(* IEC 61131-3 sources: daoli-st-library/DL_Process (part 60) *)

(* ---- FB_DL_AgvDockingHandshake.st ---- *)
(*==============================================================================
 * 组件名称 (Component)  : FB_DL_AgvDockingHandshake
 * 所属子库 (Sublibrary) : DL_Process
 * 当前版本 (Version)    : 1.0.1
 * 组件分类 (Category)   : 功能块（FUNCTION_BLOCK）· 工站模板 · 移动载体对接交接
 * 兼容性 (Platform)     : CODESYS 3.5 / TwinCAT 3 / 汇川 InoProShop / Machine Expert；
 *                         仅依赖标准库（TON / R_TRIG / F_TRIG），握手信号全部为布尔
 *                         引脚注入，块内不含任何车辆调度、导航或总线通讯细节
 * 功能描述 (Function)   : 把「到位检测 → 双侧就绪握手 → 交接放行 → 完成确认」做成带
 *                         超时与失序诊断的交接状态机，屏蔽移动载体与固定工站两侧的
 *                         信号时序差异，产出单一放行位与握手成功单拍脉冲
 * 与既有件边界 (Scope)  : 固定段之间的连续物流握手（成组上下游节拍链）由输送链路件
 *                         承担，属长连接；本件面向移动载体与固定工站的临时对接（会话
 *                         式、一次性），握手条件含「物料在位」与「双侧就绪」双约束，
 *                         语义与生命周期都不同，不可互替
 * 状态机规模 (States)   : 七态（eIdle 0 / eWaitArrive 10 / eDockConfirm 20 /
 *                         ePermitTransfer 30 / eTransferMonitor 40 / eComplete 50 /
 *                         eFault 99）；编号留 10 间隔便于插态
 * 关键算法 (Algorithm)  :
 *   ① 到位稳定：到位信号须连续两个扫描周期为真才推进，滤掉光电单拍毛刺
 *   ② 双侧就绪：两侧就绪位须同时为真且连续两拍成立，避免单拍毛刺直接放行
 *   ③ 物料一致性：进入交接监视时快照物料在位位；过程中该位由真转假且完成确认尚未
 *      到达，即判物料丢失或错位（02E2），因为这属于「该在的时候不在」
 *   ④ 完成判定：完成确认上升沿 → 置完成保持位、对接次数累加、撤放行、出握手单拍
 *   ⑤ 失序诊断：完成确认在到位或握手阶段提前到达，属非法请求序列（02E3），直接锁
 *      故障而不吞掉，否则上游误接线会被解释成「一次成功交接」
 *   ⑥ 状态停留时长：用「状态未变则计时、状态一变即清零」的单一秒表实现，供现场
 *      判读卡在哪个阶段，不额外增加引脚
 * 码位表 (Error codes)  :
 *   16#0005_01C3【信息级】超时参数越界已钳位，不置故障位
 *   16#0005_02E0【故障级】到位确认超时
 *   16#0005_02E1【故障级】握手或交接超时（两处共用，均属未在期望时间内建立期望状态）
 *   16#0005_02E2【故障级】物料在位信号丢失
 *   16#0005_02E3【故障级】非法请求序列（完成确认提前到达）
 *   16#0005_02E4【故障级】非法状态兜底
 * R32 写入点次序审计 :
 *   bTransferComplete : ① 待机启动拍清（eIdle）→ ② 交接监视完成拍置（eTransferMonitor
 *                       ，唯一置位点）。保持特性由「不再写」实现，不设第三处写点
 *   _uErrorIdInt      : ① 首扫清（段 4）→ ② 到位超时（eWaitArrive）→ ③ 握手/交接超时
 *                       （eDockConfirm 与 eTransferMonitor 各一处，同拍只命中一处）
 *                       → ④ 物料丢失（eTransferMonitor）→ ⑤ 失序（段 5）→ ⑥ 非法状态
 *                       （ELSE）→ ⑦ 复位清（eFault）
 *   _eState           : 每拍只在 CASE 分支出口单点写入；CASE 之外仅两处（段 5 失序监视、
 *                       段 6 中止与使能撤销），均在 CASE 之前，次序固定
 *   _bMatSnap         : ① 交接监视入口快照（ePermitTransfer 转出拍）→ ② 完成与复位清
 *   tElapsed          : 仅段 10 单点派生（秒表已历时），状态机内不写
 * 设计偏离登记 (Deviations) :
 *   D1 bHandshakeOk 取「握手成功」口径，在进入放行态那一拍出脉冲；规格验收向量 V1 把
 *      该脉冲写在完成确认之后叙述，二者不冲突——脉冲发生在交接放行时刻，完成确认只
 *      负责置完成保持位，头注释按状态迁移表口径落地
 *   D2 到位与双侧就绪用「连续两拍」替代「沿后与门」等价实现，效果相同（滤单拍毛刺），
 *      但不需要额外的边沿实例，拍序更易推演
 * 验收向量 (Acceptance) :
 *   V1 正常序：到位 → 双侧就绪依序为真 → 放行位为真、握手单拍、完成确认后完成保持位
 *      为真且对接次数加一
 *   V2 到位超时：超时窗 10 秒内到位信号未建立 → 码 02E0、故障态
 *   V3 物料丢失：交接监视内物料在位由真转假且完成确认为假 → 码 02E2、放行位撤
 *   V4 完成提前：到位阶段完成确认为真 → 码 02E3、直接故障态
 *   V5 统计：交接监视停留 12 秒、监视超时 30 秒 → 上一轮时长 12 秒、累计加 12 秒
 * 开源溯源 (Origin)     : 参考包装机械与批控公开手册的「会话式交接」阶段划分与双侧
 *                         就绪语义组织，只借阶段分类与参数域；状态机、快照一致性判据、
 *                         失序诊断、码位与引脚契约为本库独立设计，clean-room 不构成
 *                         衍生作品
 * 红线自检 (Redline)    : R1 零全局表与外部变量引用、零物理地址记号 ✓｜R2 零占位符 ✓
 *                         R3 纯 IEC 61131-3 加标准库 ✓｜R4 时长比较带零值旁路、计数
 *                         饱和、无数组访问 ✓｜R5 声明行中英双语同行注释 ✓｜R6 七成员
 *                         逐一有 CASE 标签且含 ELSE 兜底 ✓｜R7 三沿检测与四定时器全
 *                         部在 CASE 之外无条件刷新 ✓
 * 修订历史 (Revision)   :
 *   2026-11-15  v1.0.0  首版入库（Round 11 · C 泳道 · 工站四件套之三）
 *   2026-11-16  v1.0.1  R13 机检 R39 修复：段 5 使能撤销分支原先把 _eState 无条件
 *                       改写为 eIdle，而故障复位沿的消化位于其后 CASE 的 eFault
 *                       分支——禁用期间按下的复位沿当拍被抹掉，_bFaultLatch 与
 *                       故障码留存至操作员补按第二次复位，期间使能回升也被
 *                       「有锁存」判据挡在待机。改为 eFault 态不被禁用覆盖
 *============================================================================*)

(*------------------------------------------------------------------------------
 * 枚举: E_DL_AgvDockState（归属 FB_DL_AgvDockingHandshake，同文件发布）
 *   七态，每个成员在主状态机中均有同名 CASE 标签（R31 完备性）
 *-----------------------------------------------------------------------------*)
TYPE E_DL_AgvDockState :
(
    eIdle            := 0,  // 待机：等到位信号 / Idle, awaiting arrival signal
    eWaitArrive      := 10, // 到位确认：等到位信号稳定 / Arrival confirmation, waiting for a stable signal
    eDockConfirm     := 20, // 对接确认：等双侧就绪同时成立 / Dock confirmation, waiting for both sides ready
    ePermitTransfer  := 30, // 放行交接：单拍过渡态 / Transfer permit, a single-scan transition state
    eTransferMonitor := 40, // 交接监视：等完成确认并监视物料在位 / Transfer monitor, watching completion and material
    eComplete        := 50, // 交接完成：保持一拍后回待机 / Complete, holds one scan then returns
    eFault           := 99  // 故障锁存：仅复位沿可退 / Fault latched, only a reset edge leaves
);
END_TYPE

(*------------------------------------------------------------------------------
 * 结构体: ST_DL_AgvDockStat（归属 FB_DL_AgvDockingHandshake）
 *   跨周期统计，由调用方持有，本块只累加，掉电保持由上层负责
 *-----------------------------------------------------------------------------*)
TYPE ST_DL_AgvDockStat :
STRUCT
    nDockCount     : UDINT;                 // 累计成功对接次数 [次] [Docking counter]
    tTotalTransfer : TIME;                  // 累计交接时长 [毫秒] [Accumulated transfer time]
    tLastCycle     : TIME;                  // 上一轮交接时长 [毫秒] [Last transfer duration]
END_STRUCT
END_TYPE

FUNCTION_BLOCK FB_DL_AgvDockingHandshake
VAR_INPUT
    bEnable           : BOOL;               // 使能，FALSE 撤回全部放行位 [Enable, withdraws all permits on FALSE]
    bReset            : BOOL;               // 复位故障，上升沿受理 [Reset fault on rising edge]
    bAbort            : BOOL;               // 中止本次交接，上升沿受理，不置故障 [Abort the handshake on rising edge, no fault]
    bAgvArrived       : BOOL;               // 载体到位光电（粗定位）[-] [Carrier presence sensor]
    bAgvDockReady     : BOOL;               // 载体侧对接机构就绪 [-] [Carrier-side dock ready]
    bStationReady     : BOOL;               // 工站侧可收料或可放料 [-] [Station-side ready]
    bMaterialOnAgv    : BOOL;               // 物料在位，交接前为载侧、交接后为站侧 [-] [Material present flag]
    bTransferDone     : BOOL;               // 下游完成接收确认 [-] [Downstream receipt confirmation]
    tArriveTimeout    : TIME := T#10S;      // 到位确认超时 [毫秒]，0 表示不监控 [Arrival timeout]
    tHandshakeTimeout : TIME := T#5S;       // 双侧就绪握手超时 [毫秒]，0 表示不监控 [Handshake timeout]
    tTransferTimeout  : TIME := T#30S;      // 交接过程超时 [毫秒]，0 表示不监控 [Transfer timeout]
END_VAR
VAR_OUTPUT
    bDockLamp         : BOOL;               // 对接允许指示灯，载体可进入 [-] [Dock-permitted lamp]
    bTransferPermit   : BOOL;               // 放行交接，可放料或可接料 [-] [Transfer permit]
    bHandshakeOk      : BOOL;               // 握手成功单拍脉冲 [-] [Single pulse when handshake succeeds]
    bTransferComplete : BOOL;               // 交接完成，保持到下次启动 [Transfer complete, held until next cycle]
    eState            : E_DL_AgvDockState;  // 主状态机当前态 [-] [Current state]
    bError            : BOOL;               // 故障锁存，需复位清除 [Latched fault]
    uErrorId          : UDINT;              // 事件码或故障码，0 表示无 [Event or fault code]
    tElapsed          : TIME;               // 当前态已耗时 [毫秒]，现场判读用 [Elapsed time in current state]
END_VAR
VAR_IN_OUT
    stStat            : ST_DL_AgvDockStat;  // 跨周期统计，调用方持有 [Persistent statistics]
END_VAR
VAR
    _eState          : E_DL_AgvDockState := E_DL_AgvDockState.eIdle;  // 内部状态寄存器，唯一真值源 [Internal state register]
    _eStateIn        : E_DL_AgvDockState := E_DL_AgvDockState.eIdle;  // 上拍状态，用于识别迁移拍 [Previous state of last scan]
    _bInit           : BOOL := FALSE;       // 首扫标志，初值 FALSE，判据 NOT _bInit [First-scan flag, R19 pattern]
    _bFaultLatch     : BOOL;                // 故障级锁存，仅复位路径清 [Fault latch, reset path only]
    _uErrorIdInt     : UDINT;               // 故障级码寄存 [Fault-level code register]
    _uInfoCode       : UDINT;               // 本拍信息级码，每拍重算 [Transient info code]
    _bStateChg       : BOOL;                // 本拍发生过状态迁移，秒表清零用 [State changed this scan]
    _bArrivePrev     : BOOL;                // 上位到位信号，稳定判据用 [Arrival signal of last scan]
    _bBothReadyPrev  : BOOL;                // 上拍双侧就绪，稳定判据用 [Both-ready of last scan]
    _bMatSnap        : BOOL;                // 交接入口物料在位快照 [Material snapshot at monitor entry]
    tArriveEff       : TIME;                // 生效到位超时 [毫秒] [Effective arrival timeout]
    tHandEff         : TIME;                // 生效握手超时 [毫秒] [Effective handshake timeout]
    tTranEff         : TIME;                // 生效交接超时 [毫秒] [Effective transfer timeout]
    tMoniEff         : TIME;                // 本次交接监视时长（钳位后）[毫秒] [Clamped monitor duration]
    bArriveIn        : BOOL;                // 到位计时输入条件，先算后调 [Arrival timer input]
    bHandIn          : BOOL;                // 握手计时输入条件，先算后调 [Handshake timer input]
    bTranIn          : BOOL;                // 交接计时输入条件，先算后调 [Transfer timer input]
    fbTrigReset      : R_TRIG;              // 复位沿检测 [Reset edge detector]
    fbTrigAbort      : R_TRIG;              // 中止沿检测 [Abort edge detector]
    fbTrigDone       : R_TRIG;              // 完成确认上升沿 [Completion rising edge]
    fbTrigMateria    : F_TRIG;              // 物料在位下降沿，丢失诊断用 [Material falling edge, loss diagnosis]
    fbTmoArrive      : TON;                 // 到位确认计时 [Arrival timer]
    fbTmoHandshake   : TON;                 // 双侧就绪握手计时 [Handshake timer]
    fbTmoTransfer    : TON;                 // 交接过程计时 [Transfer timer]
    fbTmoState       : TON;                 // 状态停留秒表 [State elapsed stopwatch]
END_VAR
VAR CONSTANT
    DL_FLOAT_EPS     : REAL := 1.0E-6;      // 浮点判等容差（预留）[-] [Float comparison epsilon]
    DL_STAT_MAX      : UDINT := 16#FFFF_FFFE; // 统计计数饱和上限 [次] [Statistics saturation limit]
    DL_TMO_MAX       : TIME := T#600S;      // 超时参数域上限 [毫秒] [Timeout upper bound]
    DL_TMAX_STATE    : TIME := T#24H;       // 状态秒表量程 [毫秒] [State stopwatch range]
    DL_TIME_MAX      : TIME := T#500H;     // 累计时长饱和上限 [毫秒] [Duration saturation limit]
    DL_INFO_TMO_CLAMP: UDINT := 16#0005_01C3; // 01C3 超时参数越界已钳位【信息级】 [Info, timeout clamped]
    DL_ERR_ARRIVE    : UDINT := 16#0005_02E0; // 02E0 到位确认超时【故障级】 [Fault, arrival timeout]
    DL_ERR_HANDSHAKE : UDINT := 16#0005_02E1; // 02E1 握手或交接超时【故障级】 [Fault, handshake or transfer timeout]
    DL_ERR_MATERIAL  : UDINT := 16#0005_02E2; // 02E2 物料在位信号丢失【故障级】 [Fault, material lost]
    DL_ERR_SEQUENCE  : UDINT := 16#0005_02E3; // 02E3 非法请求序列【故障级】 [Fault, illegal request sequence]
    DL_ERR_STATE     : UDINT := 16#0005_02E4; // 02E4 非法状态兜底【故障级】 [Fault, illegal state]
END_VAR

// ==== 段 1｜单拍输出预清零（握手脉冲每拍先清零，置位点唯一） / Single-scan pulse pre-clear, single set point
bHandshakeOk := FALSE;                      // 握手单拍先清零 [Handshake pulse pre-cleared]
_uInfoCode   := 16#0000_0000;               // 信息级码每拍重算 [Info code recomputed]

// ==== 段 2｜超时参数钳位（三个超时统一钳位，零值表示不监控） / Timeout clamping, zero disables supervision
tArriveEff := tArriveTimeout;               // 到位超时先取引脚值 [Arrival timeout from pin]
IF tArriveEff > DL_TMO_MAX THEN
    tArriveEff := DL_TMO_MAX;               // 超上限钳位 [Clamped to upper bound]
    _uInfoCode := DL_INFO_TMO_CLAMP;        // 01C3 超时参数越界已钳位【信息级】 [Info, timeout clamped]
ELSIF tArriveEff < T#0S THEN
    tArriveEff := T#0S;                     // 负值归零即不监控 [Negative means disabled]
END_IF

tHandEff := tHandshakeTimeout;              // 握手超时先取引脚值 [Handshake timeout from pin]
IF tHandEff > DL_TMO_MAX THEN
    tHandEff   := DL_TMO_MAX;               // 超上限钳位 [Clamped to upper bound]
    _uInfoCode := DL_INFO_TMO_CLAMP;        // 01C3 超时参数越界已钳位【信息级】 [Info, timeout clamped]
ELSIF tHandEff < T#0S THEN
    tHandEff := T#0S;                       // 负值归零即不监控 [Negative means disabled]
END_IF

tTranEff := tTransferTimeout;               // 交接超时先取引脚值 [Transfer timeout from pin]
IF tTranEff > DL_TMO_MAX THEN
    tTranEff   := DL_TMO_MAX;               // 超上限钳位 [Clamped to upper bound]
    _uInfoCode := DL_INFO_TMO_CLAMP;        // 01C3 超时参数越界已钳位【信息级】 [Info, timeout clamped]
ELSIF tTranEff < T#0S THEN
    tTranEff := T#0S;                       // 负值归零即不监控 [Negative means disabled]
END_IF

// ==== 段 3｜沿与定时器无条件刷新（R7 红线：严禁置于 IF / CASE 分支内） / Unconditional refresh of edges and timers
fbTrigReset(CLK := bReset);                 // 复位沿 [Reset edge]
fbTrigAbort(CLK := bAbort);                 // 中止沿 [Abort edge]
fbTrigDone(CLK := bTransferDone);           // 完成确认上升沿 [Completion rising edge]
fbTrigMateria(CLK := bMaterialOnAgv);       // 物料在位下降沿 [Material falling edge]

IF (_eState = E_DL_AgvDockState.eWaitArrive) AND (tArriveEff > T#0S) THEN
    bArriveIn := TRUE;                      // 仅到位段且监控开启时计时 [Only while waiting with supervision on]
ELSE
    bArriveIn := FALSE;                     // 其余段清零 [Cleared otherwise]
END_IF
fbTmoArrive(IN := bArriveIn, PT := tArriveEff);

IF (_eState = E_DL_AgvDockState.eDockConfirm) AND (tHandEff > T#0S) THEN
    bHandIn := TRUE;                        // 仅握手段且监控开启时计时 [Only while confirming with supervision on]
ELSE
    bHandIn := FALSE;                       // 其余段清零 [Cleared otherwise]
END_IF
fbTmoHandshake(IN := bHandIn, PT := tHandEff);

IF (_eState = E_DL_AgvDockState.eTransferMonitor) AND (tTranEff > T#0S) THEN
    bTranIn := TRUE;                        // 仅交接段且监控开启时计时 [Only while monitoring with supervision on]
ELSE
    bTranIn := FALSE;                       // 其余段清零 [Cleared otherwise]
END_IF
fbTmoTransfer(IN := bTranIn, PT := tTranEff);

// 状态秒表：本拍未发生迁移才计时；迁移后的下一拍输入断一拍，已历时清零（时基由定时器内部保证）
fbTmoState(IN := (NOT _bStateChg) AND bEnable, PT := DL_TMAX_STATE);

// ==== 段 4｜首扫初始化（R19 唯一合法范式：初值 FALSE，判据 NOT，同步后置 TRUE） / First-scan initialisation with the canonical R19 pattern
IF NOT _bInit THEN
    _eState          := E_DL_AgvDockState.eIdle;  // 状态回待机 [State to idle]
    _eStateIn        := E_DL_AgvDockState.eIdle;  // 上拍状态同步 [Previous state synced]
    _bFaultLatch     := FALSE;              // 故障锁存清零 [Fault latch cleared]
    _uErrorIdInt     := 16#0000_0000;       // 故障码清零 [Fault code cleared]
    _bStateChg       := FALSE;              // 迁移标志清零 [State change flag cleared]
    _bArrivePrev     := FALSE;              // 到位上拍值清零 [Arrival previous cleared]
    _bBothReadyPrev  := FALSE;              // 双侧就绪上拍值清零 [Both-ready previous cleared]
    _bMatSnap        := FALSE;              // 物料快照清零 [Material snapshot cleared]
    bDockLamp        := FALSE;              // 指示灯灭 [Lamp off]
    bTransferPermit  := FALSE;              // 放行撤 [Permit withdrawn]
    bTransferComplete := FALSE;             // 完成保持位清 [Complete flag cleared]
    bError           := FALSE;              // 故障标志清零 [Error cleared]
    uErrorId         := 16#0000_0000;       // 事件码清零 [Error id cleared]
    tElapsed         := T#0S;               // 状态耗时清零 [Elapsed cleared]
    stStat.nDockCount     := 0;             // 对接次数清零 [Dock counter cleared]
    stStat.tTotalTransfer := T#0S;          // 累计交接时长清零 [Total transfer cleared]
    stStat.tLastCycle     := T#0S;          // 上轮时长清零 [Last cycle cleared]
    _bInit := TRUE;                         // 首扫只做一次 [Runs exactly once]
END_IF

// ==== 段 5｜全局监视：中止优先，其次失序诊断（完成确认在到位或握手阶段提前到达） / Abort first, then out-of-sequence diagnosis
IF fbTrigAbort.Q AND bEnable
AND (_eState <> E_DL_AgvDockState.eIdle)
AND (_eState <> E_DL_AgvDockState.eFault) THEN
    _bMatSnap         := FALSE;             // 快照作废（放行由出口按状态派生，不在此重复写）[Snapshot invalidated]
    _eState           := E_DL_AgvDockState.eIdle;   // 回待机，不置故障 [Back to idle, no fault]
END_IF

IF bEnable AND (NOT _bFaultLatch) AND bTransferDone
AND ((_eState = E_DL_AgvDockState.eWaitArrive) OR (_eState = E_DL_AgvDockState.eDockConfirm)) THEN
    _bFaultLatch := TRUE;                   // 失序锁存 [Sequence fault latched]
    _uErrorIdInt := DL_ERR_SEQUENCE;        // 02E3 非法请求序列【故障级】 [Fault, illegal sequence]
    _eState      := E_DL_AgvDockState.eFault;
END_IF

// ==== 段 5 之三｜使能撤销回待机（eFault 除外：复位沿的消化权归 CASE 的 eFault 分支） / Disable returns to idle, the fault state keeps its reset edge
// R39 纪律：复位沿只在发生的那一拍为真，eFault 分支是唯一清除 _bFaultLatch 与故障码
// 的出口。若本分支无条件改写 _eState，禁用期间按下的复位沿当拍被抹掉（CASE 落到 eIdle
// 分支，其判据要求 bEnable 为真，复位判据摸不到），锁存留存且二次复位才清。
// R39: the reset edge lives one scan and is only consumed inside the eFault branch, so
// the disable override must not pre-empt it, otherwise a reset pressed while disabled
// is lost and the fault latch survives until a second press.
IF (NOT bEnable) AND (_eState <> E_DL_AgvDockState.eFault) THEN
    _eState          := E_DL_AgvDockState.eIdle;   // 使能撤销回待机（放行与灯由出口派生）[Disable returns to idle]
    _bMatSnap        := FALSE;              // 快照作废 [Snapshot invalidated]
END_IF

// ==== 段 6｜主状态机（ENUM 加 CASE 加 ELSE 兜底，七成员逐一有标签） / Main state machine, every member has its own label
CASE _eState OF
    E_DL_AgvDockState.eIdle: // 待机：载体到位且使能即进入到位确认
        IF bEnable AND bAgvArrived AND (NOT _bFaultLatch) THEN
            bTransferComplete := FALSE;     // 新会话开始，清上一轮完成保持位 [Clear last completion]
            _uErrorIdInt      := 16#0000_0000;  // 启动前必无故障 [No fault before start]
            _bArrivePrev      := TRUE;      // 到位已成立，稳定判据起点 [Arrival already true]
            _bBothReadyPrev   := FALSE;     // 双侧就绪起点复位 [Both-ready starts false]
            _eState           := E_DL_AgvDockState.eWaitArrive;
        END_IF

    E_DL_AgvDockState.eWaitArrive: // 到位确认：信号连续两拍为真才推进
        IF (NOT bAgvArrived) THEN
            _eState := E_DL_AgvDockState.eIdle;   // 载体离开，回待机 [Carrier left, back to idle]
        ELSIF _bArrivePrev AND bAgvArrived THEN
            _eState := E_DL_AgvDockState.eDockConfirm;
        ELSIF fbTmoArrive.Q THEN
            _bFaultLatch := TRUE;           // 超时锁存 [Timeout latched]
            _uErrorIdInt := DL_ERR_ARRIVE;  // 02E0 到位确认超时【故障级】 [Fault, arrival timeout]
            _eState      := E_DL_AgvDockState.eFault;
        END_IF

    E_DL_AgvDockState.eDockConfirm: // 对接确认：双侧就绪同时成立且连续两拍
        IF (NOT bAgvArrived) THEN
            _eState := E_DL_AgvDockState.eIdle;   // 载体离开，回待机 [Carrier left, back to idle]
        ELSIF bAgvDockReady AND bStationReady AND _bBothReadyPrev THEN
            bHandshakeOk := TRUE;           // 握手成功单拍，本拍唯一置位点 [Sole set point of the pulse]
            _bMatSnap    := bMaterialOnAgv; // 交接前物料在位快照 [Snapshot before transfer]
            _eState      := E_DL_AgvDockState.ePermitTransfer;
        ELSIF fbTmoHandshake.Q THEN
            _bFaultLatch := TRUE;           // 超时锁存 [Timeout latched]
            _uErrorIdInt := DL_ERR_HANDSHAKE;  // 02E1 握手或交接超时【故障级】 [Fault, handshake timeout]
            _eState      := E_DL_AgvDockState.eFault;
        END_IF

    E_DL_AgvDockState.ePermitTransfer: // 放行交接：单拍过渡，把放行与监视分开便于现场观察
        _eState := E_DL_AgvDockState.eTransferMonitor;   // 放行由出口按状态派生 [Permit derived from state]

    E_DL_AgvDockState.eTransferMonitor: // 交接监视：等完成确认，同时监视物料在位
        IF fbTrigDone.Q THEN
            bTransferComplete := TRUE;      // 完成保持，本拍唯一置位点 [Sole set point of the flag]
            IF stStat.nDockCount < DL_STAT_MAX THEN
                stStat.nDockCount := stStat.nDockCount + 1;   // 对接次数饱和累加 [Dock counter, saturated]
            END_IF
            IF fbTmoTransfer.ET > tTranEff THEN
                tMoniEff := tTranEff;       // 异常值按超时上限钳位，防污染均值 [Clamp abnormal duration]
            ELSE
                tMoniEff := fbTmoTransfer.ET;
            END_IF
            stStat.tLastCycle := tMoniEff;  // 上一轮交接时长 [Last transfer duration]
            IF stStat.tTotalTransfer < DL_TIME_MAX THEN
                stStat.tTotalTransfer := stStat.tTotalTransfer + tMoniEff;  // 累计交接时长 [Total transfer accumulated]
            END_IF
            _bMatSnap := FALSE;             // 快照用毕作废 [Snapshot consumed]
            _eState   := E_DL_AgvDockState.eComplete;
        ELSIF _bMatSnap AND fbTrigMateria.Q THEN
            _bFaultLatch := TRUE;           // 物料该在时不在，锁故障 [Material lost, fault latched]
            _uErrorIdInt := DL_ERR_MATERIAL;   // 02E2 物料在位信号丢失【故障级】 [Fault, material lost]
            _eState      := E_DL_AgvDockState.eFault;
        ELSIF fbTmoTransfer.Q THEN
            _bFaultLatch := TRUE;           // 超时锁存 [Timeout latched]
            _uErrorIdInt := DL_ERR_HANDSHAKE;  // 02E1 握手或交接超时【故障级】 [Fault, transfer timeout]
            _eState      := E_DL_AgvDockState.eFault;
        END_IF

    E_DL_AgvDockState.eComplete: // 完成：保持一拍后回待机，完成保持位由 eIdle 下场会话清
        IF bAgvArrived THEN
            _bArrivePrev := TRUE;           // 载体仍在位，为下一轮预置 [Carrier still present for the next cycle]
        ELSE
            _bArrivePrev := FALSE;
        END_IF
        _eState := E_DL_AgvDockState.eIdle;

    E_DL_AgvDockState.eFault: // 故障：等复位沿，复位后清码回待机
        IF fbTrigReset.Q THEN
            _bFaultLatch := FALSE;          // 锁存解除 [Latch released]
            _uErrorIdInt := 16#0000_0000;   // 故障码清零 [Fault code cleared]
            _bMatSnap    := FALSE;          // 快照作废 [Snapshot invalidated]
            _eState      := E_DL_AgvDockState.eIdle;
        END_IF

    ELSE // 非法枚举值兜底：回安全态并锁故障（放行由出口按状态派生为假）
        _bFaultLatch    := TRUE;            // 兜底锁存 [Fallback latch]
        _uErrorIdInt    := DL_ERR_STATE;    // 02E4 非法状态兜底【故障级】 [Fault, illegal state]
        _eState         := E_DL_AgvDockState.eFault;
END_CASE

// ==== 段 7｜稳定判据与迁移寄存器更新（每次扫描末统一更新，供下一拍判稳定与秒表清零） / Stability registers updated at scan end
_bBothReadyPrev := bAgvDockReady AND bStationReady;   // 双侧就绪上拍值 [Both-ready of this scan]
IF (_eState = E_DL_AgvDockState.eWaitArrive) THEN
    _bArrivePrev := bAgvArrived;            // 到位上拍值（仅到位段跟踪）[Arrival tracked while waiting]
END_IF
_bStateChg := (_eState <> _eStateIn);       // 本拍是否迁移 [Transition happened this scan]
_eStateIn  := _eState;                      // 迁移寄存器同步 [Previous state synced]

// ==== 段 8｜出口派生（指示灯、放行、耗时均在此单点派生） / Outlets derived at a single point
bDockLamp := (_eState = E_DL_AgvDockState.eWaitArrive)
          OR (_eState = E_DL_AgvDockState.eDockConfirm);   // 对接期间指示灯亮 [Lamp on while docking]

IF (_eState = E_DL_AgvDockState.ePermitTransfer)
OR (_eState = E_DL_AgvDockState.eTransferMonitor) THEN
    bTransferPermit := TRUE;                // 交接期间放行（与状态同源，杜绝双写冲突）[Permit while transferring]
ELSE
    bTransferPermit := FALSE;
END_IF

tElapsed := fbTmoState.ET;                  // 状态停留时长 [Elapsed in current state]

eState := _eState;                          // 状态镜像 [State mirror]
bError := _bFaultLatch;                     // 故障级派生式（R21）[Fault-level derived form]
IF _bFaultLatch THEN
    uErrorId := _uErrorIdInt;               // 故障级码优先透出 [Fault code wins]
ELSE
    uErrorId := _uInfoCode;                 // 无故障时透出信息级码 [Info code otherwise]
END_IF
END_FUNCTION_BLOCK

(* ---- FB_DL_AndonCallSystem.st ---- *)
(*==============================================================================
 * 组件名称 (Component)  : FB_DL_AndonCallSystem
 * 所属子库 (Sublibrary) : DL_Process
 * 当前版本 (Version)    : 1.0.0
 * 分类     (Category)   : 人员响应工艺功能块（Function Block · 安灯呼叫系统）
 * 作者     (Author)     : Daoli Library
 * 日期     (Date)       : 2026-11-15
 * 兼容性   (Platform)   : CODESYS 3.5 / TwinCAT 3 / 汇川 InoProShop / Schneider
 *                         Machine Expert；纯 IEC 61131-3（第 3 版）语法，
 *                         仅依赖 Standard.library（TON / R_TRIG），零厂商方言
 * 功能简介 (Function)   : 车间安灯（Andon）四级呼叫系统：缺料 / 品质 / 设备 /
 *                         维修四路呼叫源，按固定优先级（维修 > 设备 > 品质 > 缺料）
 *                         做多源同拍仲裁；呼叫生命周期为「呼叫（未应答）→ 已应答
 *                         （未解除）→ 解除」三段，未应答超阈值可升级上报；应答
 *                         时长做最近值与滚动均值统计；班次清零只清统计台账，不动
 *                         激活呼叫。
 * 职责边界 (Scope)      : ① 只做「人员响应域」的状态与统计，不驱动物理灯柱：
 *                         灯色/闪频输出由既有 FB_DL_SignalTower 承载（本块仅出
 *                         级别与状态，可与之配套组合，且不依赖其实现）；
 *                         ② 与设备级状态机（如既有 FB_DL_PackMlStateMachine 的
 *                         17 态）正交：安灯描述「谁该来、来了没有」，不做设备
 *                         启停编排；③ 不做消息推送与网络上报（升级位仅作本地
 *                         输出，推送由上层 MES 接口块按位取用）。
 * 开源溯源 (Origin)     : 来源标签 andon / omac（PackML / OMAC 人员响应域开族）。
 *                         仅参考 ISA-TR88.00.02 公开规范与 OMAC 包装机工作组公开
 *                         建模惯例中「安灯四级分类（缺料/品质/设备/维修）、应答-
 *                         解除生命周期、升级上报、班次统计」的功能分类与状态域；
 *                         本块的枚举编号（数值即仲裁权重）、状态机、滚动均值算法、
 *                         引脚契约与故障码位 100% 本库独立设计，clean-room 实现，
 *                         未复制任何来源的代码行，不构成衍生作品。
 * 公约遵循 (Convention) : 0.1/R19 首扫范式（IF (NOT _bInit)）；0.2/R21 bError 显式
 *                         排除信息级码；0.5/R7 定时器与三个边沿实例主体最前部无
 *                         条件刷新；0.6/R14 计时器语义变化断输入一拍（呼叫换级时
 *                         重置升级计时）；0.7/R15 故障级锁存仅重建路径清码；
 *                         0.9 出口默认值先赋；0.14 除法防零；0.16 阈值全常量化。
 * 红线自检 (Redline)    : 全局隔离 ✓（零全局变量表引用、零外部变量声明、零物理
 *                         地址字面记号）｜命名合规 ✓（b/n/u/f/t/a/st/e/fb/i 前缀
 *                         全覆盖）｜注释完整 ✓（声明行 100% 中英双语同行注释）｜
 *                         OOP 封装 ✓（状态全私有，仅引脚与只读输出）｜周期安全 ✓
 *                         （TON / R_TRIG 均无条件刷新）｜防御编程 ✓（算术防溢出、
 *                         均值防除零、ENUM + CASE + ELSE 兜底）｜可移植性 ✓（纯
 *                         IEC 61131-3）｜终结符成对 ✓
 * 设计要点 (Key notes)  : ① 仲裁不依赖枚举数值排序：显式 IF 链按「维修 > 设备 >
 *                         品质 > 缺料」取值，枚举数值仅作对外权重标识，防止后续
 *                         插入新级别时数值序与业务序脱钩（可维护性优先）。
 *                         ② 抢占语义：eCalled / eAcked 期间更高优先级呼叫到来即
 *                         重锁，且升级计时与升级位一并重建（旧呼叫的升级计时不再
 *                         有效）；未应答即被抢占的呼叫不计入应答笔数（它不是一次
 *                         响应），只在信息级码上留痕，避免均值被「没人来」的呼叫
 *                         污染。
 *                         ③ 应答时长来源：以长周期 TON 的 ET 作为「呼叫存活时长」
 *                         计量（PT 取 24 h 上限，正常呼叫远达不到，ET 即真实
 *                         时长），避免引入累计时钟引脚；换级/新呼叫时断输入一拍
 *                         使 ET 从零重计（公约 0.6）。
 *                         ④ 滚动均值：tAckAvg += (tAckLast − tAckAvg) / 笔数。
 *                         采用增量式而非「总和 / 笔数」，避免长班次累计和溢出；
 *                         差值用 DINT 有符号运算，避免无符号下溢。
 *                         ⑤ 班次清零语义写死：只清 tAckLast / tAckAvg / uAckCount，
 *                         不清激活呼叫与升级位（现场交接班时呼叫仍需有人响应）。
 * 偏离留档 (Deviation)  : ① 规格 VAR 段 bFirstScan 改名 _bInit（公约 0.1）；
 *                         ② 规格 VAR 段 fbEscTimer 与内部计时基准拆为两支 TON
 *                         （升级计时 + 存活计时），理由见设计要点③：单个 TON 在
 *                         tEscalate = 0（不升级）时 ET 不再累加，无法同时承担
 *                         应答时长计量。
 * 故障码表 (Error codes) :
 *                         16#0005_01A0【信息级】未应答即解除（应答统计不计入）
 *                         16#0005_01A1【信息级】多源呼叫同拍或高优先级抢占重锁
 *                         16#0005_02A0【故障级】激活呼叫级别非法（内部一致性破坏）
 *                         16#0005_02A1【故障级】非法状态兜底（枚举越界）
 * 验收向量 (Acceptance) :
 *   V1 仲裁：缺料 + 设备同拍 → 激活级别为设备（优先级 2 胜 4），信息级 01A1；
 *   V2 应答统计：呼叫 30 s 后应答 → tAckLast = 30 s、uAckCount = 1、tAckAvg
 *      = 30 s；再来一次 10 s 应答 → tAckAvg = 20 s（增量均值复算）；
 *   V3 升级：tEscalate = 120 s、未应答 120 s → bEscalate 保持型置位；应答后
 *      立即复位；
 *   V4 抢占：品质呼叫 60 s 未应答，维修呼叫到来 → 级别切维修、升级计时从零
 *      重计、bEscalate 复位，uAckCount 不变（未应答不计笔数）；
 *   V5 班次清零：bShiftReset 上升沿 → tAckLast / tAckAvg / uAckCount 归零，
 *      激活呼叫与升级位保持；
 *   V6 未应答解除：eCalled 期间 bClear 上升沿 → 回 eIdle、bCallActive FALSE、
 *      信息级 01A0、uAckCount 不变。
 * 修订历史 (Revision)   :
 *   2026-11-15  v1.0.0  首版入库（Round 09 · DL_Process 安灯呼叫件）
 *============================================================================*)

(*-----------------------------------------------------------------------------
 * 调用示例 (Instance guide)：
 *   VAR fbAndon : FB_DL_AndonCallSystem; END_VAR
 *   fbAndon(bCallMat := bBtnMaterial, bCallQual := bBtnQuality,
 *           bCallDev := bBtnDevice, bCallMaint := bBtnMaintenance,
 *           bAcknowledge := bBtnAck, bClear := bBtnClear,
 *           bShiftReset := bShiftStartPulse, tEscalate := T#120S);
 *   灯柱联动：把 fbAndon.eActiveCall 映射为灯色（维修红常亮 / 设备红闪 /
 *            品质黄 / 缺料蓝），fbAndon.bEscalate 映射为蜂鸣升级。
 *   注意：bAcknowledge / bClear / bShiftReset 均为上升沿生效，长按不会重复计数。
 *----------------------------------------------------------------------------*)

(*-----------------------------------------------------------------------------
 * 常见误用与现场提示 (Field notes)：
 *   1 呼叫位是电平输入：按钮按下保持即持续呼叫，松开且呼叫未应答时呼叫仍
 *     保持（激活呼叫在状态机内锁存），不会因松手而消失——这是安灯的基本语义。
 *   2 应答后必须显式解除（bClear）才会回 eIdle：现场常见「应答了但没消灯」，
 *     属正常设计（提醒问题尚未处理完），若需自动消灯请在上层按工艺判定解除。
 *   3 升级位不改变状态机：它只是「催一下」的上报信号，不额外占用呼叫级别。
 *   4 班次清零不清激活呼叫：交接班时若仍有未处理呼叫，新班次统计从零开始但
 *     呼叫继续升级，这是有意设计。
 *   5 应答时长按「呼叫发起到按键应答」计量，不含问题实际处理时间；需要处理
 *     时长请另用维修工单系统统计。
 *----------------------------------------------------------------------------*)

(*-----------------------------------------------------------------------------
 * 枚举: E_DL_AndonLevel（归属 FB_DL_AndonCallSystem，随本文件发布）
 * 含义: 呼叫级别。数值即对外公布的仲裁权重（小者优先），状态机内部仍用显式
 *       IF 链仲裁（见设计要点①），数值仅供 HMI 排序与上位系统对照。
 *----------------------------------------------------------------------------*)
{attribute 'strict'}
{attribute 'qualified_only'}
TYPE E_DL_AndonLevel :
(
    eNone     := 0,     // 无呼叫（No call），空闲基准值 / Baseline value when no call is pending
    eMaterial := 4,     // 缺料呼叫（Material call），最低优先级 4 / Lowest priority, weight four
    eQuality  := 3,     // 品质呼叫（Quality call），优先级 3 / Priority weight three
    eDevice   := 2,     // 设备呼叫（Device call），优先级 2 / Priority weight two
    eMaint    := 1      // 维修呼叫（Maintenance call），最高优先级 1 / Highest priority, weight one
) UINT;
END_TYPE

(*-----------------------------------------------------------------------------
 * 枚举: E_DL_AndonState（归属 FB_DL_AndonCallSystem，随本文件发布）
 * 含义: 呼叫生命周期离散状态。数值步长 10 留空位，故障态 99 排序末位。
 *----------------------------------------------------------------------------*)
{attribute 'strict'}
{attribute 'qualified_only'}
TYPE E_DL_AndonState :
(
    eIdle   := 0,      // 无呼叫：等待任一呼叫源（No call, waiting for a source）
    eCalled := 10,     // 已呼叫待应答：升级计时进行中（Called, waiting for acknowledgement）
    eAcked  := 20,     // 已应答待解除：应答已记账，等待问题处理完解除（Acknowledged, waiting for the clear）
    eFault  := 99      // 内部异常：仅班次清零沿可退（Internal fault, left only by the shift reset edge）
) UINT;
END_TYPE

(*==============================================================================
 * 功能块: FB_DL_AndonCallSystem
 * 调用约定: 每个扫描周期无条件调用一次；三个事件输入均为上升沿生效。
 * 无状态泄漏: 全部状态驻留于实例私有成员，多工位各一实例，可并行。
 *============================================================================*)
FUNCTION_BLOCK FB_DL_AndonCallSystem
VAR_INPUT
    bCallMat     : BOOL;                // 缺料呼叫（Material call），优先级 4（最低） / Priority four, the lowest
    bCallQual    : BOOL;                // 品质呼叫（Quality call），优先级 3 / Priority three
    bCallDev     : BOOL;                // 设备呼叫（Device call），优先级 2 / Priority two
    bCallMaint   : BOOL;                // 维修呼叫（Maintenance call），优先级 1（最高） / Priority one, the highest
    bAcknowledge : BOOL;                // 呼叫应答（Acknowledge），上升沿对当前激活呼叫应答 / Rising edge acknowledges the active call
    bClear       : BOOL;                // 呼叫解除（Clear call），上升沿清除当前激活呼叫 / Rising edge clears the active call
    bShiftReset  : BOOL;                // 班次清零（Shift reset），上升沿清统计台账，不清激活呼叫 / Rising edge clears the statistics only
    tEscalate    : TIME := T#120S;      // 升级上报阈值（Escalation threshold）[ms]，0 = 不升级 / Zero disables escalation
END_VAR
VAR_OUTPUT
    eActiveCall  : E_DL_AndonLevel;     // 当前激活呼叫级别（Active call level），eNone = 无 / None when idle
    bCallActive  : BOOL;                // 有未应答激活呼叫（Unacknowledged call pending）/ An unacknowledged call is pending
    bAcked       : BOOL;                // 已应答未解除（Acknowledged and not yet cleared）/ Acknowledged but not yet cleared
    bEscalate    : BOOL;                // 升级上报（Escalation raised），保持型直到应答或解除 / Held until acknowledgement or clear
    tAckLast     : TIME := T#0MS;       // 最近一次应答耗时（Last acknowledgement time）[ms] / Time from call to acknowledgement [ms]
    tAckAvg      : TIME := T#0MS;       // 平均应答耗时（Average acknowledgement time）[ms]，滚动均值 / Rolling average acknowledgement time [ms]
    uAckCount    : UDINT := 0;          // 累计应答笔数（Acknowledgement count）[笔] / Number of acknowledgements
    uErrorId     : UDINT;               // 故障码（Error code），0 = 无故障，段位 16#0005_xxxx / Error code, zero means no error
END_VAR
VAR
    _eState      : E_DL_AndonState := E_DL_AndonState.eIdle; // 呼叫主状态机（Call state machine）/ Call state machine
    _bInit       : BOOL;                // 首扫完成标志（First-scan done flag），初值 FALSE / First-scan done flag, initial FALSE
    _eActive     : E_DL_AndonLevel := E_DL_AndonLevel.eNone; // 锁存的激活级别（Latched active level）/ Latched active level
    _eHighest    : E_DL_AndonLevel;     // 本拍最高优先级呼叫（Highest call level this scan）/ Highest call level in this scan
    _uCallBits   : UINT;                // 本拍呼叫源个数（Call source count this scan）[路]，0~4 / Number of active call sources, zero to four
    _tEscEff     : TIME := T#120S;      // 生效升级阈值（Effective escalation threshold）[ms] / Effective escalation threshold [ms]
    _bEscBreak   : BOOL;                // 升级计时断输入一拍（Escalation timer break），换级重置用 / One-scan break used to restart the timer
    _bEscFeed    : BOOL;                // 升级计时器输入（Escalation timer input），先算后喂 / Computed first and then fed
    _bAgeBreak   : BOOL;                // 存活计时断输入一拍（Age timer break），新呼叫重置用 / One-scan break used to restart the age timer
    _bAgeFeed    : BOOL;                // 存活计时器输入（Age timer input），先算后喂 / Computed first and then fed
    _nDeltaMs    : DINT;                // 应答耗时差值（Deviation of the sample）[ms]，有符号 / Signed deviation of the last sample [ms]
    _nStepMs     : DINT;                // 均值增量（Mean increment）[ms]，有符号 / Signed increment of the rolling mean [ms]
    _bFaultLatch : BOOL;                // 故障锁存（Fault latch），仅班次清零沿清除 / Fault latch, cleared by the shift reset edge
    _uErrInt     : UDINT;               // 故障级码寄存（Fault-level code register），锁存型 / Latched fault-level code register
    _uInfoCode   : UDINT;               // 本拍信息级码（Info code this scan），每拍重算 / Info code recomputed every scan
    _fbEscTimer  : TON;                 // 升级计时定时器（Escalation timer），主周期无条件刷新 / Refreshed unconditionally every scan
    _fbAgeTimer  : TON;                 // 呼叫存活计时定时器（Call age timer），ET 即呼叫时长 / Its elapsed time is the call age
    _fbTrigAck   : R_TRIG;              // 应答上升沿（Acknowledge rising edge）/ Acknowledge rising edge detector
    _fbTrigClear : R_TRIG;              // 解除上升沿（Clear rising edge）/ Clear rising edge detector
    _fbTrigShift : R_TRIG;              // 班次清零上升沿（Shift reset rising edge）/ Shift reset rising edge detector
END_VAR
VAR CONSTANT
    DL_AGE_LIMIT   : TIME := T#24H;     // 存活计时上限（Age timer ceiling）[ms]，正常呼叫远达不到 / Ceiling never reached by a normal call
END_VAR

// ============================================================================
// 段 1｜输出确定性默认值先赋（公约 0.9）
//      Deterministic defaults assigned before any early exit
// ============================================================================
bCallActive := FALSE;                  // 未应答呼叫标志预清零（Pending call flag pre-cleared）
bAcked      := FALSE;                  // 已应答标志预清零（Acknowledged flag pre-cleared）
bEscalate   := FALSE;                  // 升级标志预清零（Escalation flag pre-cleared）
_uInfoCode  := 0;                      // 信息级码每拍重算（Info code recomputed every scan）
_uCallBits  := 0;                      // 呼叫源计数预清零（Call source count pre-cleared）

// ============================================================================
// 段 2｜首扫初始化（R19 范式）
//      First-scan initialization following the single legal R19 predicate
// ============================================================================
IF NOT _bInit THEN
    _bInit       := TRUE;              // 置首扫完成（First-scan done）
    _eState      := E_DL_AndonState.eIdle; // 状态复位为空闲（State reset to idle）
    _eActive     := E_DL_AndonLevel.eNone; // 激活级别置无（Active level set to none）
    tAckLast     := T#0MS;             // 最近应答耗时清零（Last acknowledgement cleared）
    tAckAvg      := T#0MS;             // 平均应答耗时清零（Average acknowledgement cleared）
    uAckCount    := 0;                 // 应答笔数清零（Acknowledgement count cleared）
    _bFaultLatch := FALSE;             // 故障锁存清零（Fault latch cleared）
    _uErrInt     := 16#0000_0000;      // 故障码清零（Fault code cleared）
END_IF

// ============================================================================
// 段 3｜定时器与边沿实例无条件周期刷新（公约 0.5 / 0.6）
//      Unconditional refresh of the timers and the three edge instances
// ============================================================================
_fbTrigAck(CLK := bAcknowledge);       // 应答沿（Acknowledge edge）
_fbTrigClear(CLK := bClear);           // 解除沿（Clear edge）
_fbTrigShift(CLK := bShiftReset);      // 班次清零沿（Shift reset edge）

IF tEscalate = T#0MS THEN
    _tEscEff := T#0MS;                 // 阈值 0 = 不升级（Zero threshold disables escalation）
ELSE
    _tEscEff := tEscalate;             // 合法阈值直通（Valid threshold passed through）
END_IF

_bAgeFeed := ((_eState = E_DL_AndonState.eCalled) OR (_eState = E_DL_AndonState.eAcked)) AND (NOT _bAgeBreak); // 存活计时输入（Age timer input）
_fbAgeTimer(IN := _bAgeFeed, PT := DL_AGE_LIMIT); // 呼叫存活计时，ET 即呼叫时长（Age timing, elapsed time is the call age）
_bAgeBreak := FALSE;                   // 断输入脉冲在实例调用后自清（Break pulse self-cleared after the call）

_bEscFeed := (_eState = E_DL_AndonState.eCalled) AND (_tEscEff > T#0MS) AND (NOT _bEscBreak); // 升级计时输入（Escalation timer input）
_fbEscTimer(IN := _bEscFeed, PT := _tEscEff); // 升级计时（Escalation timing）
_bEscBreak := FALSE;                   // 断输入脉冲自清（Break pulse self-cleared）

// ============================================================================
// 段 4｜多源仲裁（显式优先级链，不依赖枚举数值序；同拍多源置信息级）
//      Source arbitration with an explicit priority chain
// ============================================================================
_eHighest := E_DL_AndonLevel.eNone;    // 默认无呼叫（Default to no call）
IF bCallMaint THEN
    _eHighest := E_DL_AndonLevel.eMaint; // 维修最高优先级（Maintenance has the highest priority）
    _uCallBits := _uCallBits + 1;      // 呼叫源计数累加（Source count incremented）
END_IF
IF bCallDev THEN
    IF _eHighest = E_DL_AndonLevel.eNone THEN
        _eHighest := E_DL_AndonLevel.eDevice; // 设备次高优先级（Device is the second priority）
    END_IF
    _uCallBits := _uCallBits + 1;      // 呼叫源计数累加（Source count incremented）
END_IF
IF bCallQual THEN
    IF _eHighest = E_DL_AndonLevel.eNone THEN
        _eHighest := E_DL_AndonLevel.eQuality; // 品质再次（Quality is the third priority）
    END_IF
    _uCallBits := _uCallBits + 1;      // 呼叫源计数累加（Source count incremented）
END_IF
IF bCallMat THEN
    IF _eHighest = E_DL_AndonLevel.eNone THEN
        _eHighest := E_DL_AndonLevel.eMaterial; // 缺料最低（Material is the lowest priority）
    END_IF
    _uCallBits := _uCallBits + 1;      // 呼叫源计数累加（Source count incremented）
END_IF

IF _uCallBits > 1 THEN
    _uInfoCode := 16#0005_01A1;        // 0005_01A1 多源呼叫同拍，按固定优先级仲裁【信息级】（Multiple sources arbitrated, info level）
END_IF

// ============================================================================
// 段 5｜班次清零（只清统计台账，不清激活呼叫；R15 顺带解除故障锁存）
//      Shift reset clears the statistics only, never the active call
// ============================================================================
IF _fbTrigShift.Q THEN
    tAckLast     := T#0MS;             // 最近应答耗时清零（Last acknowledgement cleared）
    tAckAvg      := T#0MS;             // 平均应答耗时清零（Average acknowledgement cleared）
    uAckCount    := 0;                 // 应答笔数清零（Acknowledgement count cleared）
    _bFaultLatch := FALSE;             // 班次清零同时解除内部故障锁存（The shift edge also releases the fault latch）
    _uErrInt     := 16#0000_0000;      // 故障码清零（Fault code cleared）
    IF _eState = E_DL_AndonState.eFault THEN
        _eState := E_DL_AndonState.eIdle; // 故障态经班次清零退回空闲（Fault state returns to idle）
    END_IF
END_IF

// ============================================================================
// 段 6｜内部一致性校验（激活呼叫存在但级别为无 → 内部异常）
//      Internal consistency check, an active call without a level is illegal
// ============================================================================
IF ((_eState = E_DL_AndonState.eCalled) OR (_eState = E_DL_AndonState.eAcked)) AND
   (_eActive = E_DL_AndonLevel.eNone) THEN
    _bFaultLatch := TRUE;              // 一致性破坏锁故障（Consistency break latches a fault）
    _uErrInt     := 16#0005_02A0;      // 0005_02A0 激活呼叫级别非法【故障级】（Illegal active call level, fault level）
    _eState      := E_DL_AndonState.eFault;
END_IF

// ============================================================================
// 段 7｜主状态机（ENUM + CASE + ELSE 兜底；抢占重锁 + 应答统计 + 升级）
//      Main state machine with preemption, statistics and escalation
// ============================================================================
CASE _eState OF

    E_DL_AndonState.eIdle: // 无呼叫：任一呼叫源即起呼（Idle, any source raises a call）
        IF _eHighest <> E_DL_AndonLevel.eNone THEN
            _eActive   := _eHighest;   // 锁存最高优先级级别（Latch the highest level）
            _bAgeBreak := TRUE;        // 存活计时从零重计（Age timer restarted）
            _bEscBreak := TRUE;        // 升级计时从零重计（Escalation timer restarted）
            _eState    := E_DL_AndonState.eCalled; // 进已呼叫态（Enter the called state）
        END_IF

    E_DL_AndonState.eCalled: // 已呼叫待应答（Called, waiting for acknowledgement）
        IF (_eHighest <> E_DL_AndonLevel.eNone) AND (_eHighest = E_DL_AndonLevel.eMaint) AND
           (_eActive <> E_DL_AndonLevel.eMaint) THEN
            _eActive   := E_DL_AndonLevel.eMaint; // 维修呼叫抢占一切（Maintenance preempts everything）
            _bAgeBreak := TRUE;        // 存活计时重计（Age timer restarted）
            _bEscBreak := TRUE;        // 升级计时重计，升级位随之重建（Escalation restarted, the raise bit is rebuilt）
            _uInfoCode := 16#0005_01A1; // 0005_01A1 高优先级抢占重锁【信息级】（Preemption re-lock, info level）
        ELSIF (_eHighest = E_DL_AndonLevel.eDevice) AND
              ((_eActive = E_DL_AndonLevel.eQuality) OR (_eActive = E_DL_AndonLevel.eMaterial)) THEN
            _eActive   := E_DL_AndonLevel.eDevice; // 设备抢占品质与缺料（Device preempts quality and material）
            _bAgeBreak := TRUE;        // 存活计时重计（Age timer restarted）
            _bEscBreak := TRUE;        // 升级计时重计（Escalation restarted）
            _uInfoCode := 16#0005_01A1; // 0005_01A1 高优先级抢占重锁【信息级】（Preemption re-lock, info level）
        ELSIF (_eHighest = E_DL_AndonLevel.eQuality) AND (_eActive = E_DL_AndonLevel.eMaterial) THEN
            _eActive   := E_DL_AndonLevel.eQuality; // 品质抢占缺料（Quality preempts material）
            _bAgeBreak := TRUE;        // 存活计时重计（Age timer restarted）
            _bEscBreak := TRUE;        // 升级计时重计（Escalation restarted）
            _uInfoCode := 16#0005_01A1; // 0005_01A1 高优先级抢占重锁【信息级】（Preemption re-lock, info level）
        END_IF

        IF _fbTrigAck.Q THEN
            tAckLast   := _fbAgeTimer.ET; // 应答耗时 = 呼叫存活时长（Acknowledgement time equals the call age）
            uAckCount  := uAckCount + 1;  // 应答笔数累加（Acknowledgement count incremented）
            IF uAckCount <= 1 THEN
                tAckAvg := tAckLast;      // 首笔均值等于样本（The first sample seeds the mean）
            ELSE
                _nDeltaMs := TIME_TO_DINT(tAckLast) - TIME_TO_DINT(tAckAvg); // 有符号差值，避免无符号下溢（Signed deviation avoids underflow）
                _nStepMs  := _nDeltaMs / UDINT_TO_DINT(uAckCount);           // 增量 = 差值 / 笔数（Increment is the deviation over the count）
                tAckAvg   := tAckAvg + DINT_TO_TIME(_nStepMs);               // 增量式滚动均值（Incremental rolling mean）
            END_IF
            _eState    := E_DL_AndonState.eAcked; // 进已应答态（Enter the acknowledged state）
        ELSIF _fbTrigClear.Q THEN
            _uInfoCode := 16#0005_01A0; // 0005_01A0 未应答即解除，不计应答笔数【信息级】（Cleared without an acknowledgement, info level）
            _eActive   := E_DL_AndonLevel.eNone; // 级别归无（Level cleared）
            _bAgeBreak := TRUE;        // 存活计时复位（Age timer reset）
            _bEscBreak := TRUE;        // 升级计时复位（Escalation timer reset）
            _eState    := E_DL_AndonState.eIdle; // 回空闲（Back to idle）
        END_IF

    E_DL_AndonState.eAcked: // 已应答待解除（Acknowledged, waiting for the clear）
        IF _fbTrigClear.Q THEN
            _eActive   := E_DL_AndonLevel.eNone; // 级别归无（Level cleared）
            _bAgeBreak := TRUE;        // 存活计时复位（Age timer reset）
            _bEscBreak := TRUE;        // 升级计时复位（Escalation timer reset）
            _eState    := E_DL_AndonState.eIdle; // 回空闲（Back to idle）
        ELSIF ((_eHighest = E_DL_AndonLevel.eMaint) AND (_eActive <> E_DL_AndonLevel.eMaint)) OR
              ((_eHighest = E_DL_AndonLevel.eDevice) AND
               ((_eActive = E_DL_AndonLevel.eQuality) OR (_eActive = E_DL_AndonLevel.eMaterial))) OR
              ((_eHighest = E_DL_AndonLevel.eQuality) AND (_eActive = E_DL_AndonLevel.eMaterial)) THEN
            _eActive   := _eHighest;   // 仅更高优先级重起呼叫，同级不重复触发（Only a strictly higher level re-raises）
            _bAgeBreak := TRUE;        // 新呼叫存活计时从零（New call age restarted）
            _bEscBreak := TRUE;        // 新呼叫升级计时从零（New call escalation restarted）
            _uInfoCode := 16#0005_01A1; // 0005_01A1 已应答期间更高优先级抢占【信息级】（Preemption while acknowledged, info level）
            _eState    := E_DL_AndonState.eCalled; // 回到待应答（Back to the called state）
        END_IF

    E_DL_AndonState.eFault: // 内部异常：仅班次清零沿可退（Fault, left only by the shift edge）
        _eActive := E_DL_AndonLevel.eNone; // 级别归无，输出安全（Level cleared for a safe output）
        _bEscBreak := TRUE;            // 升级计时复位（Escalation timer reset）
        _bAgeBreak := TRUE;            // 存活计时复位（Age timer reset）

    ELSE
        _bFaultLatch := TRUE;          // 非法状态兜底锁存（Illegal state latched）
        _uErrInt     := 16#0005_02A1;  // 0005_02A1 非法状态兜底【故障级】（Illegal state fallback, fault level）
        _eState      := E_DL_AndonState.eFault; // 进故障态（Enter the fault state）
END_CASE

// ============================================================================
// 段 8｜出口映射（级别、标志派生、升级判据、故障级码优先透出）
//      Outlet mapping with fault-level codes taking priority over info codes
// ============================================================================
eActiveCall := _eActive;               // 激活级别出口（Active level outlet）
bCallActive := (_eState = E_DL_AndonState.eCalled); // 未应答呼叫派生（Pending call derived form）
bAcked      := (_eState = E_DL_AndonState.eAcked);  // 已应答派生（Acknowledged derived form）
bEscalate   := (_eState = E_DL_AndonState.eCalled) AND (_tEscEff > T#0MS) AND _fbEscTimer.Q; // 升级保持型派生（Escalation derived and held）

uErrorId := _uInfoCode;                // 信息级码先透出（Info code exposed first）
IF _bFaultLatch OR (_eState = E_DL_AndonState.eFault) THEN
    uErrorId := _uErrInt;              // 故障级码优先（Fault-level code has priority）
END_IF
END_FUNCTION_BLOCK

(* ---- FB_DL_AsrsSlotAllocSeq.st ---- *)
(*==============================================================================
 * 组件名称 (Component)  : FB_DL_AsrsSlotAllocSeq
 * 所属子库 (Sublibrary) : DL_Process ｜ 版本 (Version) : 1.0.1 ｜ 2026-11-24
 * 码位     (Code Segment): 16#0005_2140（DL_Process 段内 21xx 子带，继 2100 顺排）
 * 复杂度   (Complexity) : C4
 * 兼容性   (Platform)   : CODESYS 3.5+ / TwinCAT 3 / 汇川 InoProShop / 施耐德 Machine Expert
 *                         仅依赖 IEC 61131-3 标准库（TON / R_TRIG），零厂商私有库
 * 开源溯源 (Provenance) : menes97/ayran-mini-fabrika / FB_Asrs / MIT /
 *                         借鉴点：货位分配「请求—应答」的 ack_seq / res_seq 序号同步与冲突回退语义
 *                         （未复制任何实现行，按 IEC 61131-3 重写为六相状态机 + 序号单点写入）
 * 功能描述 (Function)   : 立库货位分配与取放握手。上位下发分配请求（iReqSlot + diReqSeq），本件先做
 *                         合法性校验（入库目标必须空闲、且不能被其他任务锁闭），再进入握手相把请求
 *                         序号下发为 diOutSeq，等待对端 diAckSeq 回齐同一序号；回齐即放行（bGrant
 *                         单拍）并锁存实际分配货位。冲突（货位非空 / 应答超时）走 eRetry 净额回退，
 *                         最多 3 轮，耗尽转故障级 34。
 *                         **序号三律**：① 下发序号 _diOutSeq 全件唯一写入点（eValidate 通过相、
 *                         eRetry 回退清零点、复位点），禁止两处同拍写；② 序号超前（diAckSeq >
 *                         diOutSeq）判故障级 35——对端序号快于本端只能是对端残留或双主机，
 *                         任何「等待其自愈」的写法都是把错配隐藏成超时；③ 序号比较一律直比
 *                         `>` / `=`，不做减法防溢出假设（DINT 全值域可比，减法反而引入回绕）。
 *                         **bAllocReq 取上升沿**：电平保持不重复触发（R79 教训），重复分配必须
 *                         由上位撤请求再起，避免同一请求被连发当成多次分配。
 *                         **bEnable = FALSE 语义（R191 二选一，本件选「降级为安全值 + 置标志」）**：
 *                         放行撤销、下发序号清零、相位回 eIdle；已完成的 iAllocSlot 保留（事实不撤回）。
 * 接口     (Interface)  : 输入 bEnable / bReset（上升沿）/ bAllocReq（上升沿有效）/ iReqSlot /
 *                         diReqSeq / diAckSeq / bStoreMode / bSlotFree / bSlotLocked / tAckTimeout；
 *                         输出 eState（E_DL_AsrsSlotAllocSeq_State）/ bBusy / bDone（放行同拍单拍）/
 *                         bError / iErrCode / diOutSeq / bGrant（单拍）/ iAllocSlot / iConflictCnt。
 * 状态迁移表 (State Transition Table)：
 *   ① eIdle → eValidate：bEnable 且 rtAlloc.Q（请求上升沿）；拍 N 进入 / 本拍行为：冲突计数与
 *      信息码归零，拒绝一切放行 / 拍 N+1 转出至 eValidate。
 *   ② eValidate → eHandshake：目标货位合法（出库，或入库且空闲），且未被锁闭；拍 N 进入 /
 *      本拍行为：下发序号 _diOutSeq := diReqSeq（全件唯一写入点之一）/ 拍 N+1 转出至 eHandshake。
 *   ③ eValidate → eRetry：入库且目标货位非空；拍 N 进入 / 本拍行为：冲突计数 +1、信息级 31 /
 *      拍 N+1 转出至 eRetry。
 *   ④ eValidate → eFault：目标货位被锁闭（故障级 32）。段 7 段尾迁移闸统一迁相。
 *   ⑤ eHandshake → eCommit：diAckSeq = diOutSeq 且无锁存（本拍合法事件优先，R275）；拍 N 进入 /
 *      本拍行为：拒绝超时判定（事件已消化）/ 拍 N+1 转出至 eCommit。
 *   ⑥ eHandshake → eRetry：tonAck.Q（应答超时）；拍 N 进入 / 本拍行为：冲突计数 +1、信息级 33 /
 *      拍 N+1 转出至 eRetry。
 *   ⑦ eHandshake → eFault：diAckSeq > diOutSeq（序号超前，故障级 35）。
 *   ⑧ eRetry → eValidate：冲突计数 < 3；拍 N 进入 / 本拍行为：下发序号清零、拒绝放行 /
 *      拍 N+1 转出至 eValidate。
 *   ⑨ eRetry → eFault：冲突计数 ≥ 3（重试耗尽，故障级 34）。
 *   ⑩ eCommit → eIdle：单拍放行；拍 N 进入 / 本拍行为：bGrant 与 bDone 置单拍、iAllocSlot 锁存
 *      请求货位、拒绝重复放行 / 拍 N+1 转出至 eIdle。
 *   ⑪ eFault → eIdle：bReset 上升沿；拍 N 进入 / 本拍行为：清锁存、错误码、下发序号、冲突计数 /
 *      拍 N+1 转出至 eIdle。出口穷举、不滞留故障态。
 *   ⑫ ELSE（非法枚举值）→ eFault，码 99（R6 兜底）。
 * 边界     (Boundary)   : ① 一个 TON 与两个 R_TRIG 全部在 CASE 外无条件调用（R7）；tonAck 的 IN 含
 *                            NOT .Q 自复位项（R188），禁靠外部沿清零。
 *                         ② 序号超前判据只在 eHandshake 相内生效：eIdle 相 _diOutSeq 为 0 而
 *                            diAckSeq 可能仍为上一轮的非零值，若在空闲相判超前会误报（域证明）。
 *                         ③ eValidate 为零驻留判定相：每个分支都在本拍定相（放行 / 回退 / 故障），
 *                            不存在等待，故无需超时兜底；eCommit 为单拍放行相，同样零驻留。
 *                            eHandshake 是唯一的等待收敛相，由 tonAck（PT := _tAck）兜底（R448）。
 *                         ④ 时间参数两级回退（FB32-3）：tAckTimeout 越域（< 50ms 或 > 1h）回默认常量
 *                            T#5S，默认常量本身在有效域内，故无需二级钳定；回退不置故障（不新增码位）。
 *                         ⑤ DINT 序号比较全用 `>` / `=` 直比，不做加法/减法（无溢出路径，R4 无除法）。
 *                         ⑥ 零全局耦合（无 GVL / VAR_EXTERNAL / %I / %Q，R1 / R2）。
 * 码表     (Codes)      : 本件按派单指定使用小整数码。信息级（永不置 bError，随新请求起点重算）：
 *                         31 = 货位非空（入库目标已被占用，转回退）；反证：该场景无任何输出位变化
 *                              （bGrant 仍假、iAllocSlot 不变），仅凭输出组合不可能观测到进过 eValidate。
 *                         33 = 应答超时（对端未回齐序号，转回退）；反证：与 31 的输出组合完全同形，
 *                              两者唯一差别是成因，必须独立成码。
 *                         故障级（置 bError，锁存至 bReset 沿）：
 *                         32 = 目标货位被锁闭；反证：被锁闭时 bSlotFree 可能仍为真，与「正常放行前
 *                              拍」输出同形，只能靠码区分。
 *                         34 = 重试耗尽（冲突计数达 3）；反证：耗尽拍与普通回退拍输出全同
 *                              （iConflictCnt 已为 3 是唯一差别），且必须能被 bError 过滤上送。
 *                         35 = 序号超前（diAckSeq > diOutSeq）；反证：该场景本拍无超时、无冲突计数
 *                              变化，与「静默等待」完全同形，不报码即永久沉默。
 *                         36 = 请求序号非法（diReqSeq <= 0，未初始化禁参与握手，v1.0.1 新增）；
 *                              反证：diReqSeq=0 时 diAckSeq 初值同为 0，握手判据 (diAckSeq=_diOutSeq)
 *                              立即成立 → 零握手直接放行，输出与「正常放行拍」完全同形，只能靠码区分。
 *                              契约：diAckSeq 必须为发布后新值；提前应答或复用序号将走 33→34 耗尽（fail-closed）。
 *                         99 = 非法状态枚举值（ELSE 兜底）。
 * 分工声明 (Scope)      : 货位号有效性（1..库位总数）与货位台账维护归上游货位管理器；堆垛机行走
 *                         与取放机构归 DL_Motion 轴类件；出库货位选择策略（先进先出 / 就近）归
 *                         上层调度算法件。本件只做**一次分配事务的校验—握手—放行**时序。
 * 归属     (Ownership)  : E_DL_AsrsSlotAllocSeq_State 归属本文件（全库唯一定义，R264）。
 * 命名偏离 (Naming Ex.) : 本件按派单原文保留 i 前缀表示 INT（iReqSlot / iErrCode / iAllocSlot /
 *                         iConflictCnt），di 前缀表示 DINT（diReqSeq / diAckSeq / diOutSeq）；
 *                         与规范 1.2 节 n 前缀存在登记偏离，接口契约优先不改名。
 * 红线自检 (Redline)    : R1 ✓ 零 GVL / VAR_EXTERNAL ｜ R2 ✓ 零 %I/%Q ｜ R3 ✓ 纯 IEC 61131-3
 *                         （TON / R_TRIG）｜ R4 ✓ 无除法、无浮点、无 ABS(x-x) 判据（本件无浮点入参）
 *                         R5 ✓ 逐行同行中英双语注释 ｜ R6 ✓ 六态 ENUM + CASE + ELSE 兜底
 *                         R7 ✓ TON / R_TRIG 全在 CASE 外无条件调用 ｜ R8 ✓ 无 METHOD（全内联）
 *                         R10 ✓ 无构造式转换 ｜ R11 ✓ 声明全分号结尾 ｜ R12 ✓ ENUM 成员用 :=
 *                         R14 ✓ 无 PROPERTY ｜ R16 ✓ 不引用任何外部 FB/FC。
 * 修订历史 (Revision)   : 2026-11-24  v1.0.0  R81-B 首版
 *                          2026-11-24  v1.0.1  R81-C 补 diReqSeq<=0 闸(码36)+发布时 ack 快照，消零握手假放行（闸席 FAIL(LOGIC) 修法）
 * 验收向量 (Acceptance) :
 *   V1 入库正常：bStoreMode=TRUE、bSlotFree=TRUE、bSlotLocked=FALSE、iReqSlot=42、diReqSeq=7、
 *      diAckSeq 由 0 变 7 → eState 走 eIdle→eValidate→eHandshake→eCommit→eIdle；diOutSeq=7、
 *      bGrant 单拍为 TRUE、iAllocSlot=42、bDone 单拍为 TRUE、iErrCode=0、bError=FALSE。
 *   V2 货位非空：bStoreMode=TRUE、bSlotFree=FALSE 恒真 → 每轮 iConflictCnt+1、iErrCode=31；
 *      第 3 轮后 eState=eFault、iErrCode=34、bError=TRUE、bGrant=FALSE。
 *   V3 应答超时：diAckSeq 恒 0、tAckTimeout=T#1S → 每轮 tonAck 超时 iConflictCnt+1、iErrCode=33；
 *      第 3 轮后 eState=eFault、iErrCode=34、bError=TRUE。
 *   V4 序号超前：diReqSeq=5、diAckSeq=9 → eState=eHandshake 首拍即 eState=eFault、iErrCode=35、
 *      bError=TRUE；bReset 上升沿 → eState=eIdle、bError=FALSE、iErrCode=0、diOutSeq=0。
 *   V5 货位锁闭：bSlotLocked=TRUE → eState=eFault、iErrCode=32、bError=TRUE；bReset 上升沿可退出。
 *   V6 撤使能：eHandshake 中 bEnable=FALSE → eState=eIdle、diOutSeq=0、bGrant=FALSE、bError=FALSE。
 *============================================================================*)

(*-----------------------------------------------------------------------------
 * 枚举: E_DL_AsrsSlotAllocSeq_State（货位分配事务相位；eFault 为安全相）
 *----------------------------------------------------------------------------*)
TYPE E_DL_AsrsSlotAllocSeq_State :
(
    eIdle      := 0,    // 空闲：等分配请求上升沿 / Idle: waiting for the allocation request rising edge
    eValidate  := 10,   // 校验相：货位空闲与锁闭判定，零驻留 / Validate: slot-free and lock checks, no dwell
    eHandshake := 20,   // 握手相：下发序号并等对端回齐 / Handshake: publish the sequence and wait for the acknowledgement
    eCommit    := 30,   // 放行相：单拍输出 bGrant 并锁存货位 / Commit: one-scan grant and slot latching
    eRetry     := 40,   // 回退相：净额回退或耗尽转故障，零驻留 / Retry: net rollback or exhaustion to fault, no dwell
    eFault     := 90    // 故障安全相：锁存成因，放行撤销 / Fault safe phase: latched cause, grant withdrawn
);
END_TYPE

FUNCTION_BLOCK FB_DL_AsrsSlotAllocSeq
VAR_INPUT
    bEnable      : BOOL := FALSE;       // 使能：FALSE 撤销放行并回空闲 / Enable, FALSE withdraws the grant and returns to idle
    bReset       : BOOL := FALSE;       // 复位（上升沿，清锁存/下发序号/冲突计数）/ Reset rising edge clearing latch, output sequence and conflict count
    bAllocReq    : BOOL := FALSE;       // 分配请求（上升沿有效，电平保持不重复触发）/ Allocation request, rising edge only
    iReqSlot     : INT := 0;            // 请求货位号，有效性由上游货位管理器保证 [货位] / Requested slot number, validity guaranteed upstream
    diReqSeq     : DINT := 0;           // 请求序号（本端事务号）[序号] / Request sequence number of this transaction
    diAckSeq     : DINT := 0;           // 对端已确认序号（回齐即握手成功）[序号] / Acknowledged sequence number from the counterpart
    bStoreMode   : BOOL := TRUE;        // 作业模式：TRUE = 入库，FALSE = 出库 / Mode, TRUE for storing, FALSE for retrieving
    bSlotFree    : BOOL := FALSE;       // 目标货位空闲（入库判据）/ Target slot is free, used in store mode
    bSlotLocked  : BOOL := FALSE;       // 目标货位被其他任务锁闭（任何模式均致命）/ Target slot locked by another task, fatal in both modes
    tAckTimeout  : TIME := T#5S;        // 应答超时，有效域 50ms..1h，越域回默认 [s] / Acknowledgement timeout, out of domain falls back to the default
END_VAR
VAR_OUTPUT
    eState       : E_DL_AsrsSlotAllocSeq_State;   // 当前相位出口（段 8 单点映射）/ Current phase outlet mapped once at segment 8
    bBusy        : BOOL;                // 事务进行中（校验/握手/回退/放行）/ Transaction in progress
    bDone        : BOOL;                // 放行完成单拍脉冲 / One-scan completion pulse
    bError       : BOOL;                // 故障锁存标志 / Fault latch flag
    iErrCode     : INT := 0;            // 错误码（故障期锁存回放，非故障期为当前信息码）/ Error code, latched code in fault and the info code otherwise
    diOutSeq     : DINT := 0;           // 下发序号（对端应回齐此值）/ Published sequence number the counterpart must acknowledge
    bGrant       : BOOL;                // 放行单拍脉冲（仅 eCommit 一拍）/ One-scan grant pulse emitted only in eCommit
    iAllocSlot   : INT := 0;            // 实际分配货位（放行拍锁存，撤使能不清）/ Actually allocated slot, latched on grant and kept on disable
    iConflictCnt : INT := 0;            // 冲突累计次数，达 3 判耗尽 [次] / Conflict counter, exhaustion at three
END_VAR
VAR
    _eState      : E_DL_AsrsSlotAllocSeq_State := E_DL_AsrsSlotAllocSeq_State.eIdle;   // 内部相位（CASE 唯一写入目标）/ Internal phase, the only CASE write target
    _bFaultLatch : BOOL := FALSE;       // 故障锁存位（仅 bReset 上升沿清除）/ Fault latch bit, cleared only by the bReset rising edge
    _iErrLatch   : INT := 0;            // 锁存故障码（故障期唯一回放源，FB33-1）/ Latched fault code, the only replay source during fault
    _iInfoCode   : INT := 0;            // 信息级码（31/33，永不置 bError，新请求起点重算）/ Info-level code, never raises bError, recomputed at each new request
    _iErrTmp     : INT := 0;            // 当拍故障首因中间量 / First fault cause of this scan
    _bFaultReq   : BOOL := FALSE;       // 当拍故障请求标志（段 7 统一锁存）/ Fault request of this scan latched at segment 7
    _diOutSeq    : DINT := 0;           // 下发序号内部量（全件唯一写入点集合）/ Internal published sequence with its single-write point set
    _diAckPublish : DINT := 0;         // 下发时刻的 ack 快照，用于拦截陈旧 ack 二次放行（v1.0.1）/ Ack snapshot at publish time, blocks stale-ack re-grant
    _bGrantPulse : BOOL := FALSE;       // 放行内部单拍位（段 1 预置，段 8 映射）/ Internal one-scan grant bit preset at segment 1
    _bDonePulse  : BOOL := FALSE;       // 完成内部单拍位（段 1 预置，段 8 映射）/ Internal one-scan done bit preset at segment 1
    _iAllocSlot  : INT := 0;            // 内部实际货位（放行拍锁存）/ Internal allocated slot latched on the grant scan
    _iConflictCnt : INT := 0;           // 内部冲突计数 [次] / Internal conflict counter
    _tAck        : TIME := T#5S;        // 应答超时钳定值（两级回退结果）[s] / Clamped acknowledgement timeout after the two-level fallback
    rtReset      : R_TRIG;              // bReset 边沿实例（段 3 无条件调用，R18）/ bReset edge instance called unconditionally
    rtAlloc      : R_TRIG;              // bAllocReq 边沿实例（段 3 无条件调用，防电平重复触发）/ bAllocReq edge instance preventing level retriggering
    tonAck       : TON;                 // 应答超时计时器（段 3 无条件调用）/ Acknowledgement timeout timer called unconditionally
END_VAR
VAR CONSTANT
    DL_ASA_RETRY_MAX : INT := 3;                 // 冲突回退上限，达此判耗尽 [次] / Conflict retry limit, exhaustion at this count
    DL_ASA_CNT_ZERO  : INT := 0;                 // 计数零基准 [-] / Zero base for counters
    DL_ASA_ONE       : INT := 1;                 // 整数一（计数步进）[1] / Integer one used for stepping
    DL_ASA_T_MIN     : TIME := T#50MS;           // 应答超时下限 [s] / Acknowledgement timeout lower bound
    DL_ASA_T_MAX     : TIME := T#1H;             // 应答超时上限 [s] / Acknowledgement timeout upper bound
    DL_ASA_ACK_DEF   : TIME := T#5S;             // 应答超时默认回退值（本身在有效域内）[s] / Default fallback timeout, already inside the valid domain
END_VAR

(* —— 段 1：中间量预置（只清单拍标志与扫描量，不清序号 / 冲突计数 / 锁存，FB32-1） —— *)
_iErrTmp     := 0;                        // 当拍故障首因复位 / Scan first fault cause reset
_bFaultReq   := FALSE;                    // 当拍故障请求复位 / Scan fault request reset
_bGrantPulse := FALSE;                    // 放行单拍位预置（单拍路径唯一预置点，FB51-8）/ Grant pulse preset, the single preset point
_bDonePulse  := FALSE;                    // 完成单拍位预置（单拍路径唯一预置点，FB51-8）/ Done pulse preset, the single preset point

(* —— 段 2：时间参数两级回退（越域回默认常量，默认常量在域内故无需二级钳定，FB32-3） —— *)
IF (tAckTimeout < DL_ASA_T_MIN) OR (tAckTimeout > DL_ASA_T_MAX) THEN
    _tAck := DL_ASA_ACK_DEF;              // 越域：回一级默认常量 / Out of domain: fall back to the default constant
ELSE
    _tAck := tAckTimeout;                 // 域内：原值采用 / Inside the domain: take the value as given
END_IF

(* —— 段 3：边沿与定时器（CASE 外无条件调用，R7；IN 含 NOT .Q 自复位，R188） —— *)
rtReset(CLK := bReset);                   // bReset 边沿无条件刷新（R18）/ bReset edge refreshed unconditionally
rtAlloc(CLK := bAllocReq);                // 分配请求边沿无条件刷新（防电平重复触发，R79）/ Allocation request edge refreshed unconditionally
tonAck(IN := (_eState = E_DL_AsrsSlotAllocSeq_State.eHandshake) AND (NOT tonAck.Q) AND (NOT _bFaultLatch),
       PT := _tAck);                      // 应答超时计时（仅握手相，自复位后逐轮回退再起）/ Acknowledgement timeout running only in the handshake phase

(* —— 段 4：状态机主体（唯一相位写入点；故障只置请求，锁存与迁相由段 7 执行，R21） —— *)
CASE _eState OF
    E_DL_AsrsSlotAllocSeq_State.eIdle :
        (* 迁移①：请求上升沿且使能 → 校验相；拍 N 进入 / 本拍行为：冲突计数与信息码归零 / 拍 N+1 转出 *)
        IF bEnable AND rtAlloc.Q THEN
            _iConflictCnt := DL_ASA_CNT_ZERO;                         // 新请求起点：冲突计数归零 / New request: conflict counter cleared
            _iInfoCode    := 0;                                       // 新请求起点：信息码归零 / New request: info code cleared
            _eState       := E_DL_AsrsSlotAllocSeq_State.eValidate;   // 进校验相 / Move to validate
        END_IF

    E_DL_AsrsSlotAllocSeq_State.eValidate :
        (* 零驻留判定相：三个分支都在本拍定相，无等待故无超时兜底需求（边界③） *)
        IF diReqSeq <= 0 THEN
            _iErrTmp   := 36;                                     // 故障级：请求序号非法（0/负=未初始化，禁参与握手）/ Fault: illegal request sequence
            _bFaultReq := TRUE;                                   // 请求段 7 锁存 / Request the latch at segment 7
        ELSIF bSlotLocked THEN
            _iErrTmp   := 32;                                     // 故障级：目标货位被锁闭 / Fault: target slot locked
            _bFaultReq := TRUE;                                   // 请求段 7 锁存 / Request the latch at segment 7
        ELSIF bStoreMode AND (NOT bSlotFree) THEN
            _iConflictCnt := _iConflictCnt + DL_ASA_ONE;           // 入库目标非空：冲突净额 +1 / Store target occupied: one net conflict
            _iInfoCode    := 31;                                   // 信息级：货位非空（不置 bError）/ Info: slot not free, bError stays false
            _eState       := E_DL_AsrsSlotAllocSeq_State.eRetry;   // 迁移③：转回退 / Move to retry
        ELSE
            _diOutSeq := diReqSeq;                                 // 下发序号写入点①：请求序号下发（唯一写入点集合）/ Write point one: publish the request sequence
            _diAckPublish := diAckSeq;                             // v1.0.1：记录发布时刻 ack 快照 / v1.0.1: snapshot ack at publish time
            _eState   := E_DL_AsrsSlotAllocSeq_State.eHandshake;   // 迁移②：进握手相 / Move to handshake
        END_IF

    E_DL_AsrsSlotAllocSeq_State.eHandshake :
        (* 同拍竞态处理：本拍合法事件（序号回齐）优先于超时迁移（R275），超时判定列最后 *)
        IF (diAckSeq = _diOutSeq) AND (diAckSeq <> _diAckPublish) AND (NOT _bFaultLatch) THEN
            (* v1.0.1 修法：同序号陈旧 ack 不得二次放行（fail-closed）/ v1.0.1: a stale equal ack must not re-grant *)
            _eState := E_DL_AsrsSlotAllocSeq_State.eCommit;         // 迁移⑤：回齐且无锁存，进放行相（R274 全量复检）/ Acknowledged, move to commit
        ELSIF diAckSeq > _diOutSeq THEN
            _iErrTmp   := 35;                                       // 故障级：序号超前（对端快于本端）/ Fault: sequence ahead of the published value
            _bFaultReq := TRUE;                                     // 请求段 7 锁存 / Request the latch at segment 7
        ELSIF tonAck.Q THEN
            _iConflictCnt := _iConflictCnt + DL_ASA_ONE;            // 应答超时：冲突净额 +1 / Acknowledgement timeout: one net conflict
            _iInfoCode    := 33;                                    // 信息级：应答超时（不置 bError）/ Info: acknowledgement timeout, bError stays false
            _eState       := E_DL_AsrsSlotAllocSeq_State.eRetry;    // 迁移⑥：转回退 / Move to retry
        END_IF

    E_DL_AsrsSlotAllocSeq_State.eRetry :
        (* 拍 N 进入（冲突发生）/ 本拍行为：耗尽判或净额回退并清下发序号 / 拍 N+1 转出（R80 三段式） *)
        IF _iConflictCnt >= DL_ASA_RETRY_MAX THEN
            _iErrTmp   := 34;                                       // 故障级：重试耗尽 / Fault: retries exhausted
            _bFaultReq := TRUE;                                     // 请求段 7 锁存 / Request the latch at segment 7
        ELSE
            _diOutSeq := 0;                                         // 下发序号写入点②：回退清零点（单赋值，禁两处同拍写）/ Write point two: rollback clearing
            _eState   := E_DL_AsrsSlotAllocSeq_State.eValidate;     // 迁移⑧：回校验相 / Back to validate
        END_IF

    E_DL_AsrsSlotAllocSeq_State.eCommit :
        (* 迁移⑩：放行单拍；拍 N 进入 / 本拍行为：bGrant 与 bDone 各置一次、货位锁存、拒绝重复放行 / 拍 N+1 转出至 eIdle *)
        IF NOT _bFaultLatch THEN
            _iAllocSlot  := iReqSlot;                               // 实际分配货位锁存 / Allocated slot latched
            _bGrantPulse := TRUE;                                   // 放行内部单拍置位（段 8 映射）/ Internal grant pulse raised and mapped at segment 8
            _bDonePulse  := TRUE;                                   // 完成内部单拍置位（段 8 映射）/ Internal done pulse raised and mapped at segment 8
            _eState      := E_DL_AsrsSlotAllocSeq_State.eIdle;      // 迁移⑩：回空闲相 / Back to idle
        END_IF

    E_DL_AsrsSlotAllocSeq_State.eFault :
        (* 迁移⑪：复位沿出口（唯一出口，穷举可达）/ 拍 N 进入 / 本拍行为：清锁存与序号，放行由段 8 归假 / 拍 N+1 转出至 eIdle *)
        IF rtReset.Q THEN
            _bFaultLatch  := FALSE;                                 // 清故障锁存 / Clear the fault latch
            _iErrLatch    := 0;                                     // 清锁存故障码 / Clear the latched fault code
            _iInfoCode    := 0;                                     // 清信息码 / Clear the info code
            _diOutSeq     := 0;                                     // 下发序号写入点③：复位清零点 / Write point three: reset clearing
            _iConflictCnt := DL_ASA_CNT_ZERO;                       // 冲突计数清零 / Conflict counter cleared
            _eState       := E_DL_AsrsSlotAllocSeq_State.eIdle;     // 回空闲相，不滞留故障态 / Back to idle, never parked in fault
        END_IF

ELSE
    (* 迁移⑫：非法枚举兜底（R6） *)
    IF NOT _bFaultLatch THEN
        _iErrLatch   := 99;                    // 故障级：非法状态枚举值 / Fault: illegal state enum value
        _bFaultLatch := TRUE;                  // 置故障锁存（码位赋值 3 行内配对，R45）/ Latch the fault within three lines
    END_IF
END_CASE

(* —— 段 7：当拍故障请求锁存 + 段尾故障迁移闸 + 撤使能降级（R191 已声明为降级+置标志） —— *)
IF _bFaultReq AND (NOT _bFaultLatch) THEN
    _iErrLatch   := _iErrTmp;                  // 锁存当拍首因 / Latch the first cause of this scan
    _bFaultLatch := TRUE;                      // 置故障锁存 / Latch the fault
END_IF
IF _bFaultLatch AND (_eState <> E_DL_AsrsSlotAllocSeq_State.eFault) THEN
    _eState := E_DL_AsrsSlotAllocSeq_State.eFault;   // 锁存即迁相（段尾统一执行，FB50-1④）/ Latch forces the fault phase at the tail
END_IF
IF (NOT bEnable) AND (NOT _bFaultLatch) AND (_eState <> E_DL_AsrsSlotAllocSeq_State.eIdle) THEN
    _diOutSeq    := 0;                         // 撤使能：撤销下发序号（握手作废）/ Disable: published sequence withdrawn
    _bGrantPulse := FALSE;                     // 撤使能：放行撤销 / Disable: grant withdrawn
    _eState      := E_DL_AsrsSlotAllocSeq_State.eIdle;   // 撤使能：回空闲相 / Disable: back to idle
END_IF

(* —— 段 8：统一出口（单点映射，禁在 CASE 后无条件清零 CASE 内赋值标识符，FB33-1） —— *)
eState       := _eState;                       // 相位映射 / Phase mapping
bBusy        := (_eState = E_DL_AsrsSlotAllocSeq_State.eValidate)
                OR (_eState = E_DL_AsrsSlotAllocSeq_State.eHandshake)
                OR (_eState = E_DL_AsrsSlotAllocSeq_State.eRetry)
                OR (_eState = E_DL_AsrsSlotAllocSeq_State.eCommit);   // 事务进行中 / Transaction in progress
bGrant       := _bGrantPulse AND (NOT _bFaultLatch);   // 放行输出（故障期强制撤销）/ Grant output forced off during fault
bDone        := _bDonePulse AND (NOT _bFaultLatch);    // 完成输出（故障期强制撤销）/ Done output forced off during fault
bError       := _bFaultLatch;                  // 故障标志取锁存位 / Fault flag taken from the latch
IF _bFaultLatch THEN
    iErrCode := _iErrLatch;                    // 故障期回放锁存码（FB33-1）/ Replay the latched code during fault
ELSE
    iErrCode := _iInfoCode;                    // 非故障期输出信息码（31/33 永不置 bError，R101）/ Info code outside fault, never raising bError
END_IF
diOutSeq     := _diOutSeq;                     // 下发序号映射 / Published sequence mapping
iAllocSlot   := _iAllocSlot;                   // 实际货位映射（撤使能保留事实，不撤回）/ Allocated slot mapping, kept on disable
iConflictCnt := _iConflictCnt;                 // 冲突计数映射 / Conflict counter mapping
END_FUNCTION_BLOCK
